// TIA Portal V20 export
// export: Created 2026-10-12T05:42:33.9214397Z, ExportSetting WithDefaults, DisplayName Totally Integrated Automation Portal, DisplayVersion V20, DisplayName TIA Portal Openness, DisplayVersion V20, DisplayName TIA Portal Teamcenter Gateway, DisplayVersion V20, DisplayName TIA Portal Version Control Interface, DisplayVersion V20, DisplayName SINAMICS Startdrive Advanced, DisplayVersion V20 SP1 Update 2, DisplayName SINAMICS Startdrive G110M, G120, G120C, G120D, G120P, G115D, DisplayVersion V20 SP1 Update 2, DisplayName SINAMICS Startdrive G130, G150, S120, S150, SINAMICS MV, G220, S200, S210, DisplayVersion V20 SP1 Update 2, DisplayName STEP 7 Professional, DisplayVersion V20, DisplayName STEP 7 Safety, DisplayVersion V20, DisplayName WinCC Basic/Comfort/Advanced, DisplayVersion V20, DisplayName WinCC Professional, DisplayVersion V20, DisplayName WinCC Unified, DisplayVersion V20
FUNCTION "FRK_CfgRestore_PressDemoUnit" : Void   // FC174, SCL
{ S7_Optimized_Access := 'TRUE' }
VERSION : 0.1
// stored: AutoNumber true, IsIECCheckEnabled false, SetENOAutomatically false, UDAEnableTagReadback false
   VAR_IN_OUT
      Core : "FRK_Core";
      Status : "ST_ModuleStatus";
      StationCfg : "ST_PressDemoStationCfg";
      ConfigStageStationCfg : "ST_PressDemoStationCfg";
      ConfigDefaultStationCfg : "ST_PressDemoStationCfg";
   END_VAR
   VAR_TEMP
      RootIndex : Int;
      Ok : Bool;
      Stored : Bool;
   END_VAR
BEGIN

   #RootIndex := "FRK_ConfigRoot"(RegIndex := #Core.RegIndex);
   IF #RootIndex = 0 THEN
       RETURN;
   END_IF;
   #Ok := TRUE;
   #ConfigStageStationCfg := #ConfigDefaultStationCfg;
   "FRK_CfgDef_PressDemoUnit"(FieldIndex := 1);
   IF "FRK_ConfigFind"(Scope := #Status.Name, Key := "FRK_ConfigScratch".Entry.WriteKey, ModelCode := '') = 0 THEN
       IF #ConfigDefaultStationCfg.RequireTwoHandStart THEN
           "FRK_ConfigScratch".Entry.ValueText := WSTRING#'true';
       ELSE
           "FRK_ConfigScratch".Entry.ValueText := WSTRING#'false';
       END_IF;
       #Stored := "FRK_ConfigPut"(Scope := #Status.Name, ModelCode := '', Text := "FRK_ConfigScratch".Entry.ValueText, RootIndex := #RootIndex);
       IF NOT "FRK_ConfigRuntime".Fresh THEN
           #Ok := FALSE;
           "FRK_ConfigLoss"(RootIndex := #RootIndex,
                            Scope := #Status.Name);
       END_IF;
   END_IF;
   #Stored := "FRK_ConfigGet"(Scope := #Status.Name, ModelCode := '');
   #Ok := #Ok AND #Stored;
   IF #Stored THEN
       #ConfigStageStationCfg.RequireTwoHandStart := "FRK_ConfigScratch".Value.Flag;
   END_IF;
   "FRK_CfgDef_PressDemoUnit"(FieldIndex := 2);
   IF "FRK_ConfigFind"(Scope := #Status.Name, Key := "FRK_ConfigScratch".Entry.WriteKey, ModelCode := '') = 0 THEN
       "FRK_ConfigScratch".Entry.ValueText := DINT_TO_WSTRING(TIME_TO_DINT(#ConfigDefaultStationCfg.TransferSettleTime));
       #Stored := "FRK_ConfigPut"(Scope := #Status.Name, ModelCode := '', Text := "FRK_ConfigScratch".Entry.ValueText, RootIndex := #RootIndex);
       IF NOT "FRK_ConfigRuntime".Fresh THEN
           #Ok := FALSE;
           "FRK_ConfigLoss"(RootIndex := #RootIndex,
                            Scope := #Status.Name);
       END_IF;
   END_IF;
   #Stored := "FRK_ConfigGet"(Scope := #Status.Name, ModelCode := '');
   #Ok := #Ok AND #Stored;
   IF #Stored THEN
       #ConfigStageStationCfg.TransferSettleTime := DINT_TO_TIME(LINT_TO_DINT("FRK_ConfigScratch".Value.Number));
   END_IF;
   "FRK_CfgDef_PressDemoUnit"(FieldIndex := 3);
   IF "FRK_ConfigFind"(Scope := #Status.Name, Key := "FRK_ConfigScratch".Entry.WriteKey, ModelCode := '') = 0 THEN
       "FRK_ConfigScratch".Entry.ValueText := DINT_TO_WSTRING(TIME_TO_DINT(#ConfigDefaultStationCfg.PressSettleTime));
       #Stored := "FRK_ConfigPut"(Scope := #Status.Name, ModelCode := '', Text := "FRK_ConfigScratch".Entry.ValueText, RootIndex := #RootIndex);
       IF NOT "FRK_ConfigRuntime".Fresh THEN
           #Ok := FALSE;
           "FRK_ConfigLoss"(RootIndex := #RootIndex,
                            Scope := #Status.Name);
       END_IF;
   END_IF;
   #Stored := "FRK_ConfigGet"(Scope := #Status.Name, ModelCode := '');
   #Ok := #Ok AND #Stored;
   IF #Stored THEN
       #ConfigStageStationCfg.PressSettleTime := DINT_TO_TIME(LINT_TO_DINT("FRK_ConfigScratch".Value.Number));
   END_IF;
   IF #Ok THEN
       #StationCfg := #ConfigStageStationCfg;
   ELSE
       #StationCfg := #ConfigDefaultStationCfg;
       "FRK_ConfigLoss"(RootIndex := #RootIndex,
                        Scope := #Status.Name);
       "FRK_CfgDef_PressDemoUnit"(FieldIndex := 1);
       IF #ConfigDefaultStationCfg.RequireTwoHandStart THEN
           "FRK_ConfigScratch".Entry.ValueText := WSTRING#'true';
       ELSE
           "FRK_ConfigScratch".Entry.ValueText := WSTRING#'false';
       END_IF;
       #Stored := "FRK_ConfigPut"(Scope := #Status.Name, ModelCode := '', Text := "FRK_ConfigScratch".Entry.ValueText, RootIndex := #RootIndex);
       "FRK_CfgDef_PressDemoUnit"(FieldIndex := 2);
       "FRK_ConfigScratch".Entry.ValueText := DINT_TO_WSTRING(TIME_TO_DINT(#ConfigDefaultStationCfg.TransferSettleTime));
       #Stored := "FRK_ConfigPut"(Scope := #Status.Name, ModelCode := '', Text := "FRK_ConfigScratch".Entry.ValueText, RootIndex := #RootIndex);
       "FRK_CfgDef_PressDemoUnit"(FieldIndex := 3);
       "FRK_ConfigScratch".Entry.ValueText := DINT_TO_WSTRING(TIME_TO_DINT(#ConfigDefaultStationCfg.PressSettleTime));
       #Stored := "FRK_ConfigPut"(Scope := #Status.Name, ModelCode := '', Text := "FRK_ConfigScratch".Entry.ValueText, RootIndex := #RootIndex);
   END_IF;
END_FUNCTION
